(* IEC 61131-3 sources: Lasal-MCP/examples/SampleSource/LASALScreenAdvancedSolution/LASALScreenAdvancedSolution/LASALScreenAdvacnedSolution/Stations/Terminal/HMI/Network, 1 file *)

(* ---- ConfigObjects.st ---- *)
FUNCTION GLOBAL TAB TASK_CONF
_K_TASK, _K_REAL,
_K_END_VAR,

_K_TASK, _K_CYCLIC,
_K_END_VAR,

_K_TASK, _K_BACKGROUND,
_K_END_VAR,

_K_END_CONF
END_FUNCTION

FUNCTION GLOBAL TAB IPR_CONF
_K_IPR
	0$UINT,
_K_END_VAR,
_K_END_CONF
END_FUNCTION

FUNCTION GLOBAL TAB CONFIG_TABLES
00086$UINT,
0$UINT, 0, 11, "_ALARMDISPLAY",
0$UINT, 0, 11, "_ALARMX0PARA",
0$UINT, 0, 2, "_ALARMX1PARA",
0$UINT, 0, 21, "_ALARMXBUFFER",
0$UINT, 0, 1, "_BIT32",
0$UINT, 0, 1, "_BIT32RAM",
0$UINT, 0, 4, "_CAN",
0$UINT, 1, 4, "_CHECKONLINESTATUS",
0$UINT, 1, 0, "_CHECKSUM",
0$UINT, 1, 20, "_FILESYS",
0$UINT, 0, 15, "_GLOBAL",
0$UINT, 1, 3, "_GRAFIX",
0$UINT, 0, 1, "_HOTALARM",
0$UINT, 0, 5, "_LANGUAGESELECTION",
0$UINT, 0, 2, "_LIMITMAX",
0$UINT, 0, 2, "_LIMITMIN",
0$UINT, 0, 126, "_LSE",
0$UINT, 1, 1, "_MULTITASK",
0$UINT, 0, 3, "_MYIO",
0$UINT, 0, 5, "_OSKERNEL",
0$UINT, 0, 6, "_OSZILSE",
0$UINT, 0, 0, "_OSZILSEBACKGROUND",
0$UINT, 0, 1, "_RADIO32",
0$UINT, 0, 1, "_RADIO32RAM",
0$UINT, 0, 3, "_SCREEN",
0$UINT, 0, 15, "_SCROLLAREA",
0$UINT, 0, 8, "_SCROLLAREA2",
0$UINT, 0, 0, "_STDLIB",
0$UINT, 2, 1, "_SYNCTIMEHMI",
0$UINT, 0, 9, "_SYSDATETIME",
0$UINT, 0, 0, "_SYSMSG",
0$UINT, 1, 1, "_TASKOBJECTCONTROL",
0$UINT, 1, 1, "_TOOLCAT",
0$UINT, 0, 1, "_XACCESS",
0$UINT, 1, 8, "ALARMDISPLAYLIST",
0$UINT, 1, 2, "ALARMTITLELINE",
0$UINT, 0, 0, "CIRLEMYIO",
0$UINT, 0, 4, "CRITICALSECTION",
0$UINT, 1, 1, "DATAMANAGER",
0$UINT, 1, 1, "DATAMANAGERFIFO",
0$UINT, 1, 0, "DATAMANAGERPRIORITY",
0$UINT, 0, 0, "DATARECORD",
0$UINT, 0, 0, "DATARECORDSAVE",
0$UINT, 0, 1, "DATASERVICECLIENT",
0$UINT, 1, 37, "DISPLAYSETTINGS",
0$UINT, 0, 0, "FILEHANDLING",
0$UINT, 0, 0, "FILEREAD",
0$UINT, 0, 10, "GETBROADCASTDATA",
0$UINT, 0, 2, "GETTASKHANDLE",
0$UINT, 0, 1, "GRAPHIC",
0$UINT, 0, 0, "INDICATOR",
0$UINT, 0, 0, "INPUTMYIO",
0$UINT, 2, 0, "KEYPADANUMSTDTEMPLATE",
0$UINT, 2, 0, "KEYPADIMAGESSTDTEMPLATE",
0$UINT, 1, 0, "KEYPADNUMSTDTEMPLATE",
0$UINT, 1, 22, "MERKEREX",
0$UINT, 0, 0, "MYCAROUSEL",
0$UINT, 0, 0, "MYCOLORBAR",
0$UINT, 0, 0, "MYFIRSTMYIO",
0$UINT, 0, 0, "MYHEADER",
0$UINT, 0, 0, "MYKEYBOARDCODE",
0$UINT, 0, 0, "MYRECALCULATE",
0$UINT, 0, 0, "MYSCROLLLIST",
0$UINT, 0, 0, "MYUSERCALL",
0$UINT, 0, 0, "MYVALUES",
0$UINT, 1, 0, "PRELOADINGSCREENS",
0$UINT, 1, 18, "PROJECTGLOBAL",
0$UINT, 1, 3, "RAM",
0$UINT, 1, 17, "RAMEX",
0$UINT, 1, 1, "RAMRINGBUFFER",
0$UINT, 1, 13, "SCREENSAVER",
0$UINT, 0, 34, "SIGCLIB",
0$UINT, 1, 11, "STRING",
0$UINT, 1, 84, "STRINGINTERNAL",
0$UINT, 1, 10, "STRINGRAM",
0$UINT, 0, 1, "SYSTEM",
0$UINT, 1, 5, "SYSTEMLOGGING",
0$UINT, 1, 19, "TCPCOMMUNICATION",
0$UINT, 1, 0, "TCPCOMMUNICATIONLOGFILTER",
0$UINT, 1, 4, "TCPCOMMUNICATIONLOGVIEWER",
0$UINT, 1, 3, "TITLELINE",
0$UINT, 1, 4, "TOUCHCALIB",
0$UINT, 1, 13, "USB_DATAEXCHANGE",
0$UINT, 1, 6, "USBDETECTION",
0$UINT, 0, 0, "USEIMAGESCHEME",
0$UINT, 1, 3, "VIRTUALBASEINIT",
ONE_CFG$UINT, 0, 0, "ONE_CarouselNet",
ONE_CFG$UINT, 0, 0, "ONE_ExamplesNet",
ONE_CFG$UINT, 0, 0, "ONE_GlobalNet",
ONE_CFG$UINT, 0, 0, "ONE_LseRtkAlarm",
ONE_CFG$UINT, 0, 0, "ONE_LseRtkMain",
ONE_CFG$UINT, 0, 0, "ONE_MyIONet",
ONE_CFG$UINT, 1, 0, "ONE_NewAgeAlarmVis",
ONE_CFG$UINT, 1, 0, "ONE_NewAgeSettings",
ONE_CFG$UINT, 0, 0, "ONE_ScrollNet",
ONE_CFG$UINT, 1, 0, "ONE_STDCommunicationToPLC",
ONE_CFG$UINT, 2, 0, "ONE_STDSettingsHMI",
ONE_CFG$UINT, 0, 0, "ONE_ValueNet",
TASK_CFG$UINT, 0, 0, "TASK_CONF",
IPR_CFG$UINT, 0, 0, "IPR_CONF",
PRJ_CFG$UINT, 0, 0, "HMI",
END_FUNCTION

#ifdef __LSLLDR_MULTIMASTER__
FUNCTION GLOBAL TAB CONFIG_MULTIMASTER
0000$UINT, 0001$UINT,
"MachineControl",
0002$UINT,
TO_UDINT(619908241), "SyncTimePLC.SyncDate", 0$USINT, 103$UINT, (0)$UDINT,
TO_UDINT(3791233966), "SyncTimePLC.SyncTime", 0$USINT, 103$UINT, (0)$UDINT,
END_FUNCTION
#endif

FUNCTION GLOBAL TAB CH_REDIRECT_EMB_TAB
0000$UINT,
00009$UINT,
"ALARMDISPLAYLIST;ALATXTLONG", "\ALARMTXTLONG.DATA",
"ALARMDISPLAYLIST;ALATXTSHORT", "\ALARMTXTSHORT.DATA",
"FILEHANDLING;DRIVENAME1", "\DRIVENAME.DATA",
"FILEHANDLING;FILEEXTENSION1", "\FILEEXTENSION.DATA",
"FILEHANDLING;FILENAME1", "\FILENAME.DATA",
"MYCAROUSEL;LASALOBJECTNAME", "\LASALOBJNAME.DATA",
"MYCAROUSEL;LSEOBJECTNAME", "\LSEOBJNAME.DATA",
"TCPCOMMUNICATION;TASKNAME", "\THREADNAME.DATA",
"USBDETECTION;DRIVELETTER", "\USBDRIVELETTER.DATA",
END_FUNCTION
